(* PLC project zarechnaya.project, CODESYS CODESYS V3.5 SP17 Patch 3 *)
(* stored: creationDateTime 2026-10-20T05:42:22.250194, modificationDateTime 1601-01-01T03:00:00 *)

(* PRG_PumpInterlock — взаимная блокировка насосов II подъёма (LD, PROGRAM: параллели, двойная катушка). Поведение (модель scenarios/reference/model_PRG_PumpInterlock.py), сети по порядку: 1. xP1Run := (xP1Ready AND NOT xP2Run) OR xP1Force; 2. xP2Run := (xP2Ready AND NOT xP1Run) OR xP2Force — читает уже новое xP1Run этого цикла; 3. xAnyRun := xP1Run OR xP2Run; 4. xAlarm := xP1Run AND xP2Run; 5. xAlarm := xEmergency — двойная катушка: последняя сеть побеждает (C2S7-GFX-DOUBLECOIL). *)
PROGRAM PRG_PumpInterlock
  VAR_INPUT
    xP1Ready : BOOL;
    xP2Ready : BOOL;
    xP1Force : BOOL;
    xP2Force : BOOL;
    xEmergency : BOOL;
  END_VAR
  VAR_OUTPUT
    xP1Run : BOOL;
    xP2Run : BOOL;
    xAnyRun : BOOL;
    xAlarm : BOOL;
  END_VAR

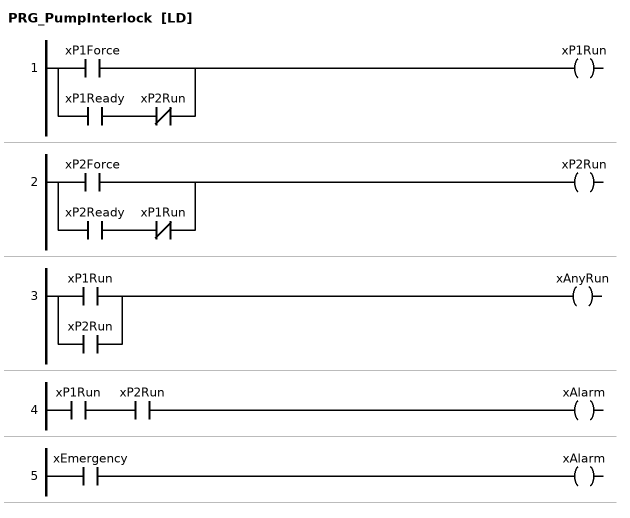
(* LD diagram, written out as Structured Text *)
(* --- network: Насос 1 --- *)
xP1Run := xP1Ready AND NOT xP2Run OR xP1Force;
(* --- network: Насос 2 --- *)
xP2Run := xP2Ready AND NOT xP1Run OR xP2Force;
(* --- network: Любой в работе --- *)
xAnyRun := xP1Run OR xP2Run;
(* --- network: Оба в работе --- *)
xAlarm := xP1Run AND xP2Run;
(* --- network: Аварийная кнопка --- *)
xAlarm := xEmergency;
END_PROGRAM
